(* IEC 61131-3 sources: avi-aoi-management/scripts/ai-eval/ngau-nhien/kho/st-tt4-trung-binh-truot/khung/src, 1 file *)

(* ---- TrungBinhTruot.st ---- *)
FUNCTION_BLOCK TrungBinhTruot
VAR_INPUT
    MAU : REAL;
    LAY_MAU : BOOL;
    RESET : BOOL;
END_VAR
VAR_OUTPUT
    TB : REAL;
    SO_MAU : INT;
    HOP_LE : BOOL;
END_VAR
    (* TODO: cài đặt theo đề bài *)
    TB := 0.0;
END_FUNCTION_BLOCK
